// TIA Portal V21 export
FUNCTION_BLOCK "Demo"   // FB10, LAD
{ S7_Optimized_Access := 'TRUE' }
   VAR_INPUT
      Start : Bool;   // Start button
   END_VAR
   VAR DB_SPECIFIC
      Ins_Delay : TON_TIME;
   END_VAR
   VAR
      Pos : Struct
         X : Int := 5;
      END_STRUCT;
   END_VAR
BEGIN

REGION Network 1: Delay
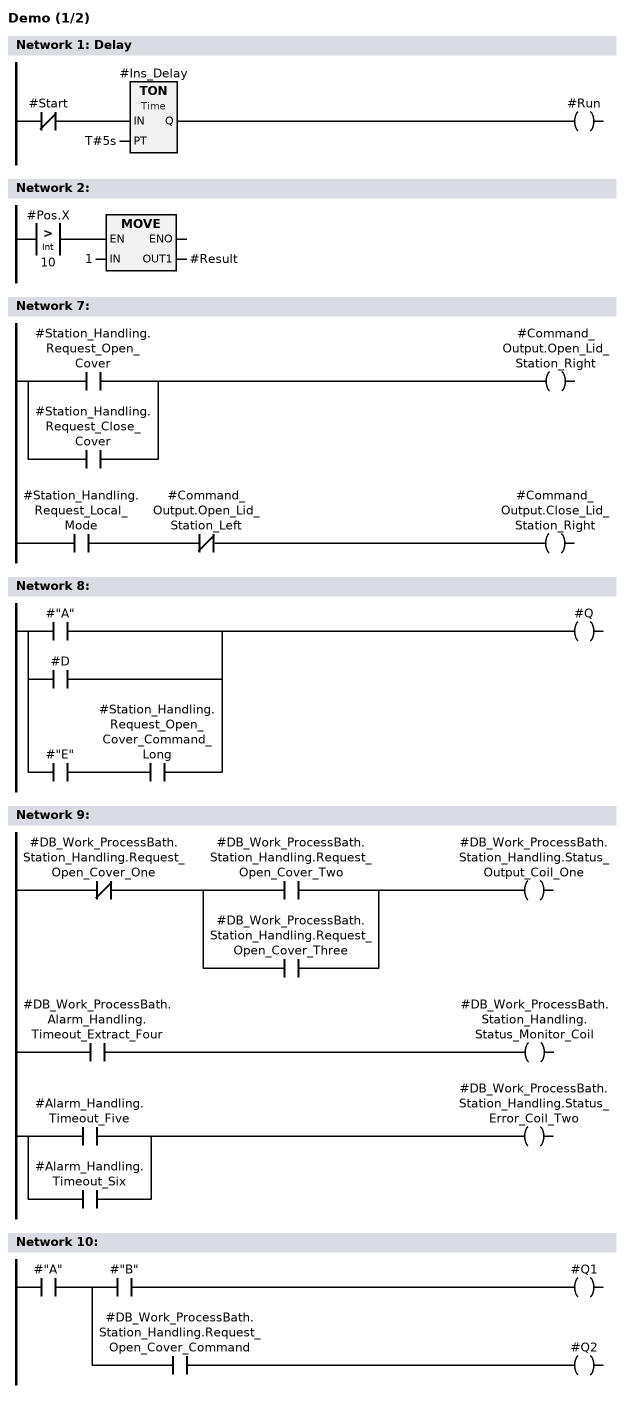
   RUNG wire#powerrail
      I_Contact( #Start )
      { S7_Templates := "time_type := Time" } #Ins_Delay.TON(pt := T#5s)
      Coil( #Run )
   END_RUNG
   // the same network as SCL:
   #Ins_Delay(in := NOT #Start, pt := T#5s);   // TON
   #Run := #Ins_Delay.q;
END_REGION

REGION Network 2
   RUNG wire#powerrail
      { S7_Templates := "SrcType := Int" } GT_Contact(in1 := #Pos.X, in2 := 10)
      Move(in := 1, out1 => #Result)
   END_RUNG
   // the same network as SCL:
   IF #Pos.X > 10 THEN #Result := 1; END_IF;
END_REGION

NETWORK
TITLE = 
      A     #Start;
      =     #Run;

REGION Network 4 (SCL)
   #Run := #Start;
   // done
END_REGION

REGION Network 6 (SCL)
   #Ins_Cfg(i_A  := "M_IBN_0", // TODO a
       io_DB  := "DB_Work".Bath[#tBathIndex]);
END_REGION

REGION Network 7
   RUNG wire#powerrail
      Contact( #Station_Handling.Request_Open_Cover )
      wire#w1
      Coil( #Command_Output.Open_Lid_Station_Right )
   END_RUNG
   RUNG wire#powerrail
      Contact( #Station_Handling.Request_Close_Cover )
   END_RUNG wire#w1
   RUNG wire#powerrail
      Contact( #Station_Handling.Request_Local_Mode )
      I_Contact( #Command_Output.Open_Lid_Station_Left )
      Coil( #Command_Output.Close_Lid_Station_Right )
   END_RUNG
   // the same network as SCL:
   #Command_Output.Open_Lid_Station_Right := #Station_Handling.Request_Open_Cover OR #Station_Handling.Request_Close_Cover;
   #Command_Output.Close_Lid_Station_Right := #Station_Handling.Request_Local_Mode AND NOT #Command_Output.Open_Lid_Station_Left;
END_REGION

REGION Network 8
   RUNG wire#powerrail
      Contact( #"A" )
      wire#w1
      Coil( #Q )
   END_RUNG
   RUNG wire#powerrail
      Contact( #D )
   END_RUNG wire#w1
   RUNG wire#powerrail
      Contact( #"E" )
      Contact( #Station_Handling.Request_Open_Cover_Command_Long )
   END_RUNG wire#w1
   // the same network as SCL:
   #Q := #"A" OR #D OR (#"E" AND #Station_Handling.Request_Open_Cover_Command_Long);
END_REGION

REGION Network 9
   RUNG wire#powerrail
      I_Contact( #DB_Work_ProcessBath.Station_Handling.Request_Open_Cover_One )
      wire#w1
      Contact( #DB_Work_ProcessBath.Station_Handling.Request_Open_Cover_Two )
      wire#w2
      Coil( #DB_Work_ProcessBath.Station_Handling.Status_Output_Coil_One )
   END_RUNG
   RUNG wire#w1
      Contact( #DB_Work_ProcessBath.Station_Handling.Request_Open_Cover_Three )
   END_RUNG wire#w2
   RUNG wire#powerrail
      Contact( #DB_Work_ProcessBath.Alarm_Handling.Timeout_Extract_Four )
      Coil( #DB_Work_ProcessBath.Station_Handling.Status_Monitor_Coil )
   END_RUNG
   RUNG wire#powerrail
      Contact( #Alarm_Handling.Timeout_Five )
      wire#w3
      Coil( #DB_Work_ProcessBath.Station_Handling.Status_Error_Coil_Two )
   END_RUNG
   RUNG wire#powerrail
      Contact( #Alarm_Handling.Timeout_Six )
   END_RUNG wire#w3
   // the same network as SCL:
   #DB_Work_ProcessBath.Station_Handling.Status_Output_Coil_One := NOT #DB_Work_ProcessBath.Station_Handling.Request_Open_Cover_One AND (#DB_Work_ProcessBath.Station_Handling.Request_Open_Cover_Two OR #DB_Work_ProcessBath.Station_Handling.Request_Open_Cover_Three);
   #DB_Work_ProcessBath.Station_Handling.Status_Monitor_Coil := #DB_Work_ProcessBath.Alarm_Handling.Timeout_Extract_Four;
   #DB_Work_ProcessBath.Station_Handling.Status_Error_Coil_Two := #Alarm_Handling.Timeout_Five OR #Alarm_Handling.Timeout_Six;
END_REGION

REGION Network 10
   #Q1 := #"A" AND #"B";
   #Q2 := #"A" AND #DB_Work_ProcessBath.Station_Handling.Request_Open_Cover_Command;
END_REGION

REGION Network 11
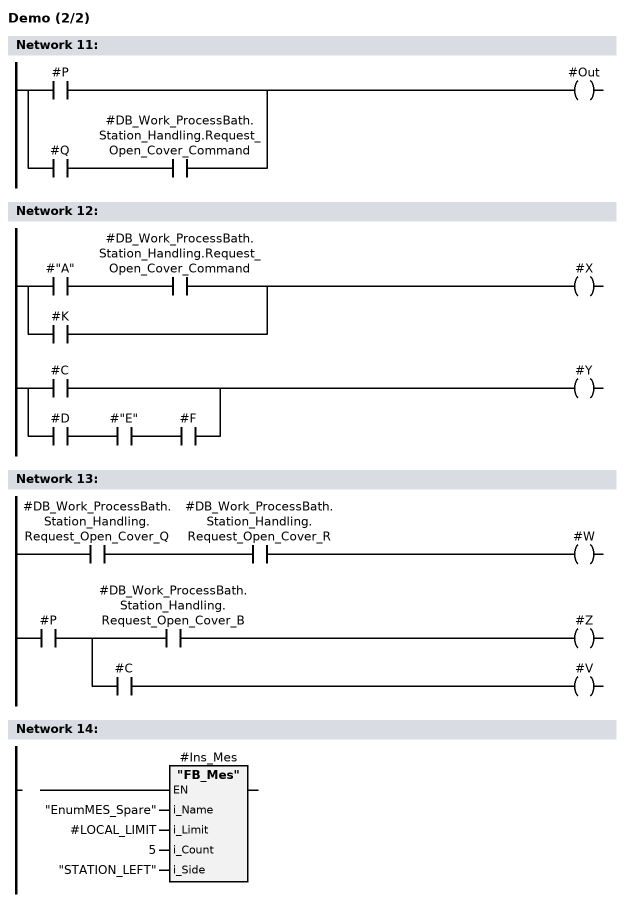
   RUNG wire#powerrail
      Contact( #P )
      wire#w1
      Coil( #Out )
   END_RUNG
   RUNG wire#powerrail
      Contact( #Q )
      Contact( #DB_Work_ProcessBath.Station_Handling.Request_Open_Cover_Command )
   END_RUNG wire#w1
   // the same network as SCL:
   #Out := #P OR (#Q AND #DB_Work_ProcessBath.Station_Handling.Request_Open_Cover_Command);
END_REGION

REGION Network 12
   #X := (#"A" AND #DB_Work_ProcessBath.Station_Handling.Request_Open_Cover_Command) OR #K;
   #Y := #C OR (#D AND #"E" AND #F);
END_REGION

REGION Network 13
   #W := #DB_Work_ProcessBath.Station_Handling.Request_Open_Cover_Q AND #DB_Work_ProcessBath.Station_Handling.Request_Open_Cover_R;
   #Z := #P AND #DB_Work_ProcessBath.Station_Handling.Request_Open_Cover_B;
   #V := #P AND #C;
END_REGION

REGION Network 14
   #Ins_Mes(i_Name := "EnumMES_Spare", i_Limit := #LOCAL_LIMIT, i_Count := 5, i_Side := "STATION_LEFT");   // "FB_Mes"
END_REGION

REGION Network 15 (SCL)
   #Ver := "GLOBAL_MAJOR";
END_REGION
END_FUNCTION_BLOCK
